(*
+------------------------+------------+----------+----------+
| Header row, column 1   | Header 2   | Header 3 | Header 4 |
| (header rows optional) |            |          |          |
+========================+============+==========+==========+
| body row 1, column 1   | column 2   | column 3 | column 4 |
+------------------------+------------+----------+----------+
| body row 2             | Cells may span columns.          |
+------------------------+------------+---------------------+
| body row 3             | Cells may  | - Table cells       |
+------------------------+ span rows. | - contain           |
| body row 4             |            | - body elements.    |
+------------------------+------------+---------------------+
*)

FUNCTION_BLOCK FB_Libdoc_GridTable
VAR_INPUT
    nVarA : INT;
    nVarB : INT;
END_VAR
VAR_OUTPUT
    nSum : INT;
END_VAR
VAR
END_VAR

END_FUNCTION_BLOCK

(* stored: Version 1.1.0.1, ProductVersion 3.1.4022.17
   POU FB_Libdoc_GridTable: Id {cbd16f47-0180-4101-957a-85db98b5fa2b}, SpecialFunc None *)
